(* PLC project Vn_fn_len, Beckhoff Automation GmbH TwinCAT PLC Control 3.5.13.21 *)
(* stored: creationDateTime 1970-01-01T00:00:00 *)

PROGRAM Vn_fn_len

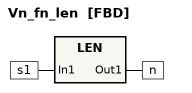
(* FBD diagram, written out as Structured Text *)
n := LEN(s1);
END_PROGRAM
